Fanuc KAREL source: KD00002.KL

PROGRAM KD00002
%NOLOCKGROUP
%CMOS2SHADOW
VAR
  I: INTEGER
  J: INTEGER
  B: BOOLEAN
  R: REAL
  S: STRING[80]
BEGIN
  I = 1
END KD00002
